(* IEC 61131-3 sources: moqui-plc/codesys-v4/moqui-plc.fbsdev/moqui.iecapp^/moqui/runtime/component/mantle-hvac/src/main/mantle/hvac, 3 files *)

(* ---- Main.fb.st ---- *)
(*
 * NOTE: In general, the Main component implements the control logic of automated industrial systems (Finite State Machine - FSM)
 * using hierarchical control architectures. It separates control policies from implementation mechanisms,
 * and diagnostic mechanisms from failure/error reaction and system reset policies.
*)

(* Example of a supervisor FSM for a civil HVAC air-handling unit (AHU).
 *
 * Topology:
 *   Mode A Thermostat cooling -> Cooling
 *   Mode B Cooling with RH% dehumidification -> Cooling  (rhControlEnabled=TRUE)
 *   Mode C Winter heating -> Heating
 *   Mode D Heating with RH% control -> Heating (rhControlEnabled=TRUE)
 *   Mode E Interval dehumidification (on/off) -> Drying
 *   Mode F Dehumidification by RH% target -> Drying (rhControlEnabled=TRUE)
 *
 * Output function - which device groups are enabled per state:
 *
 *   State          Cold Group   Hot Group   AHU Fan   Air Flow
 *   -
 *   Standby            OFF         OFF        OFF       OFF
 *   Ventilation        OFF         OFF        ON        ON
 *   Cooling            ON          OFF        ON        ON
 *   Heating            OFF         ON         ON        ON
 *   Drying             ON          ON         ON        ON
 *   Fault              OFF         OFF        OFF       OFF
 *
 * MainRuleEngine generates transition requests; Main consumes them.
 * DeviceManager orchestrates the individual device FBs.
 *
 * Call order in the PLC task:
 *   InputSignalUpdate -> Main -> DeviceManager -> OutputSignalUpdate
 *)
FUNCTION_BLOCK Main

	VAR_INPUT
		operationType : OperatingMode;
		enable : BOOL;
		deviceConfigContextResetRequest : BOOL := FALSE;
	END_VAR
	VAR_OUTPUT
		done : BOOL;
		error : BOOL;
	END_VAR
	VAR CONSTANT
		componentName : STRING := 'HVAC_DEMO_PLC';
	END_VAR
	VAR
		(* Logger facade *)
		logger : LoggerFacade;
		(* FSM transition logic *)
		ruleEngine : MainRuleEngine;
		(* Define a nested FSMs for managing air distribution subsystem. *)
		airDistribCtrl : AirDistributionController;
		(* HAL manager *)
		deviceManager : DeviceManager;
		(* Periodic logical-parameter logger *)
		logParameters : ParameterLogger;
		(* Previous status, so that the FSM state is logged on change only *)
		statusOld : MainStatus := MainStatus.Standby;
	END_VAR

	(* Logger facade init *)
	logger.enable := TRUE; logger.loggerName := componentName;

	IF NOT enable THEN RETURN; END_IF

	(* Init: device setup and configuration *)
	IF (operationType = operatingMode.Init) THEN
		logger(message := 'Setup and configuration of all devices.', level := LogLevel.DEBUG);
		(*
	     * The static device configuration parameters are mapped directly by the device config manager (recipe manager),
		 * while only the dynamic parameters are mapped below in the standby status.
		 *)
		(* Reset signal manager *)
		ec.dev.signalMgmt(operationType := SignalMgmtOperatingMode.Reset, loggerName := componentName);
		ec.dev.status := MainStatus.Standby;
		ec.dev.actualRuntime := 0;
		ec.dev.actualBreakDuration := 0;
		ec.dev.processActualDuration := 0;
		ec.dev.processRemainingDuration := 0;
		ec.dev.timeBreakEnabled := FALSE;
		ec.dev.isCompleted := FALSE;
		airDistribCtrl(operationType := OperatingMode.Init, enable := FALSE, clock1s := FALSE);
		done := FALSE;
	ELSIF deviceConfigContextResetRequest THEN
		logger(message := 'Reset HVAC device config context.', level := LogLevel.DEBUG);
		(*
	     * Lightweight reset between recipes: keep device init/homing in the Init path,
		 * but clear runtime state inherited from the previous device config.
	     *)
		ec.dev.status := MainStatus.Standby;
		ec.dev.lastStatus := MainStatus.Standby;
		ec.dev.actualRuntime := 0;
		ec.dev.actualBreakDuration := 0;
		ec.dev.processActualDuration := 0;
		ec.dev.processRemainingDuration := 0;
		ec.dev.timeBreakEnabled := FALSE;
		ec.dev.isCompleted := FALSE;
		airDistribCtrl(operationType := OperatingMode.Init, enable := FALSE, clock1s := FALSE);
		done := FALSE;
	ELSE
		(* FSM transition-condition rule engine *)
		ruleEngine(operationType := operationType);
	END_IF;

		(*
		 * Preserve the originating phase while idling in Standby so thermostat-driven
		 * Heating/Cooling recipes can stop/start repeatedly until isCompleted becomes TRUE.
		 * Init still stamps Standby, which keeps fresh-start logic for a newly loaded recipe.
		 * A temporary thermal override of Drying (Drying -> Cooling/Heating) keeps Drying as the
		 * originating phase: MainRuleEngine returns to Drying from Cooling/Heating while
		 * lastStatus = Drying, so it must stay Drying for the whole override, not for one scan.
	     *)
		IF operationType = OperatingMode.Init THEN
			ec.dev.lastStatus := ec.dev.status;
		ELSIF (ec.dev.status <> MainStatus.Standby)
				AND NOT ((ec.dev.lastStatus = MainStatus.Drying)
					AND ((ec.dev.status = MainStatus.Cooling) OR (ec.dev.status = MainStatus.Heating))) THEN
			ec.dev.lastStatus := ec.dev.status;
		END_IF;

	(* Fault overrides any other state *)
	IF ec.dev.faultRequest THEN ec.dev.status := MainStatus.Fault; END_IF;

	(* Main FSM - Output function + State-update function *)
	CASE ec.dev.status OF
	    (* Standby / Homing: all groups off, wait for the next phase request. *)
		MainStatus.Standby :
			ec.dev.standbyRequest := FALSE;

			(* FSM Output function - everything disabled *)
			ec.dev.coldGroupEnableRequest := FALSE;
			ec.dev.coldGroupDisableRequest := TRUE;
			ec.dev.hotGroupEnableRequest := FALSE;
			ec.dev.hotGroupDisableRequest := TRUE;
			ec.dev.ahuFanEnableRequest := FALSE;
			ec.dev.airFlowEnableRequest := FALSE;
			ec.dev.airFlowDisableRequest := TRUE;

			(* FSM status update function *)
			IF ec.dev.ventilationRequest THEN
				ec.dev.status := MainStatus.Ventilation;
			ELSIF ec.dev.coolingRequest THEN
				ec.dev.status := MainStatus.Cooling;
			ELSIF ec.dev.heatingRequest THEN
				ec.dev.status := MainStatus.Heating;
			ELSIF ec.dev.dryingRequest THEN
				ec.dev.status := MainStatus.Drying;
			END_IF;

	    (* Ventilation: AHU + air flow control only - no temperature conditioning. *)
		MainStatus.Ventilation :
			ec.dev.ventilationRequest := FALSE;

			(* FSM output function *)
			ec.dev.coldGroupEnableRequest := FALSE;
			ec.dev.coldGroupDisableRequest := TRUE;
			ec.dev.hotGroupEnableRequest := FALSE;
			ec.dev.hotGroupDisableRequest := TRUE;
			ec.dev.ahuFanEnableRequest := TRUE;
			ec.dev.airFlowEnableRequest := TRUE;
			ec.dev.airFlowDisableRequest := FALSE;

			(* FSM status update function *)
			IF ec.dev.standbyRequest THEN
				ec.dev.status := MainStatus.Standby;
			ELSIF ec.dev.coolingRequest THEN
				ec.dev.status := MainStatus.Cooling;
			ELSIF ec.dev.heatingRequest THEN
				ec.dev.status := MainStatus.Heating;
			ELSIF ec.dev.dryingRequest THEN
				ec.dev.status := MainStatus.Drying;
			END_IF;

	    (*
	     * Cooling: cold group + AHU + air flow control.
	     * Mode A (no RH ctrl) and Mode B (with RH dehumidification, rhControlEnabled=TRUE).
	     * In Mode B the hot group is also enabled to re-heat after dehumidification;
	     * that secondary enable is issued by MainRuleEngine via heatingRequest/dryingRequest
	     * transitions rather than here, keeping output function clean.
	     *)
		MainStatus.Cooling :
			ec.dev.coolingRequest := FALSE;

			(* FSM output function *)
			ec.dev.coldGroupEnableRequest := TRUE;
			ec.dev.coldGroupDisableRequest := FALSE;
			ec.dev.hotGroupEnableRequest := FALSE;
			ec.dev.hotGroupDisableRequest := TRUE;
			ec.dev.ahuFanEnableRequest := TRUE;
			ec.dev.airFlowEnableRequest := TRUE;
			ec.dev.airFlowDisableRequest := FALSE;

			(* FSM status update function *)
			IF ec.dev.standbyRequest THEN
				ec.dev.status := MainStatus.Standby;
			ELSIF ec.dev.dryingRequest THEN
				ec.dev.status := MainStatus.Drying;
			ELSIF ec.dev.ventilationRequest THEN
				ec.dev.status := MainStatus.Ventilation;
			END_IF;

	    (*
	     * Heating: hot group + AHU + air flow control.
	     * Mode C (no RH ctrl) and Mode D (with RH ctrl).
	     *)
		MainStatus.Heating :
			ec.dev.heatingRequest := FALSE;

			(* FSM output function *)
			ec.dev.coldGroupEnableRequest := FALSE;
			ec.dev.coldGroupDisableRequest := TRUE;
			ec.dev.hotGroupEnableRequest := TRUE;
			ec.dev.hotGroupDisableRequest := FALSE;
			ec.dev.ahuFanEnableRequest := TRUE;
			ec.dev.airFlowEnableRequest := TRUE;
			ec.dev.airFlowDisableRequest := FALSE;

			(* FSM status update function *)
			IF ec.dev.standbyRequest THEN
				ec.dev.status := MainStatus.Standby;
			ELSIF ec.dev.dryingRequest THEN
				ec.dev.status := MainStatus.Drying;
			ELSIF ec.dev.ventilationRequest THEN
				ec.dev.status := MainStatus.Ventilation;
			END_IF;

	    (*
	     * Drying: cold + hot + AHU + air flow control.
	     * Mode E (interval on/off) and Mode F (RH% controlled).
	     * During break the rule engine transitions to Standby; returns here
	     * when the break is complete.
	     *)
		MainStatus.Drying :
			ec.dev.dryingRequest := FALSE;

			(* FSM output function *)
			ec.dev.coldGroupEnableRequest := TRUE;
			ec.dev.coldGroupDisableRequest := FALSE;
			ec.dev.hotGroupEnableRequest := TRUE;
			ec.dev.hotGroupDisableRequest := FALSE;
			ec.dev.ahuFanEnableRequest := TRUE;
			ec.dev.airFlowEnableRequest := TRUE;
			ec.dev.airFlowDisableRequest := FALSE;

			(* FSM status update function *)
			IF ec.dev.standbyRequest THEN
				ec.dev.status := MainStatus.Standby;
			ELSIF ec.dev.heatingRequest THEN
				ec.dev.status := MainStatus.Heating;
			ELSIF ec.dev.coolingRequest THEN
				ec.dev.status := MainStatus.Cooling;
			ELSIF ec.dev.ventilationRequest THEN
				ec.dev.status := MainStatus.Ventilation;
			END_IF;

	    (* Fault: all groups off; wait for signal manager to clear all alarms. *)
		MainStatus.Fault :
			ec.dev.faultRequest := FALSE;

			(* FSM output function *)
			error := TRUE;
			ec.dev.coldGroupEnableRequest := FALSE;
			ec.dev.coldGroupDisableRequest := TRUE;
			ec.dev.hotGroupEnableRequest := FALSE;
			ec.dev.hotGroupDisableRequest := TRUE;
			ec.dev.ahuFanEnableRequest := FALSE;
			ec.dev.airFlowEnableRequest := FALSE;
			ec.dev.airFlowDisableRequest := TRUE;

			(* Return to Standby only when all alarms have been cleared *)
			IF (ec.dev.signalMgmt.cumulativeOutputAction = SignalOutputAction.None) THEN
				error := FALSE;
				ec.dev.status := MainStatus.Standby;
			END_IF;
	END_CASE;

	(*
	 * Air distribution is a subordinate subsystem:
	 * it runs only when the main FSM requests air flow and the recipe explicitly
	 * enables alternating high/low air distribution.
	 *)
	airDistribCtrl(
		operationType := operationType,
		enable := ec.dev.airFlowEnableRequest AND ec.dev.airDistributionEnabled,
		clock1s := ec.clks.clock1s);

	done := ec.dev.isCompleted;

	(* Log the FSM state on change only: a message every scan would fill the log buffer. *)
	IF ec.dev.status <> statusOld THEN
		CASE ec.dev.status OF
			MainStatus.Standby : logger(message := 'Standby.', level := LogLevel.Info);
			MainStatus.Ventilation : logger(message := 'Ventilation.', level := LogLevel.Info);
			MainStatus.Cooling : logger(message := 'Cooling.', level := LogLevel.Info);
			MainStatus.Heating : logger(message := 'Heating.', level := LogLevel.Info);
			MainStatus.Drying : logger(message := 'Drying.', level := LogLevel.Info);
			MainStatus.Fault : logger(message := 'Fault.', level := LogLevel.Error);
		END_CASE;
		statusOld := ec.dev.status;
	END_IF;

	(* Device orchestration (HAL) *)
	deviceManager(operationType := operationType);

	(* Log the coherent post-device-update parameter snapshot. *)
	logParameters(operationType := operationType);
	END_FUNCTION_BLOCK

(* ---- MainRuleEngine.fb.st ---- *)
(*
 * MainRuleEngine - transition-condition logic for the HVAC supervisor FSM.
 *
 * Responsibilities:
 *   1. Reset transition requests to safe defaults.
 *   2. Run the signal management engine (fault / alarm / warning detection).
 *   3. Compute boolean predicates from sensor feedback and recipe setpoints.
 *   4. Implement the per-state transition-condition rules.
 *
 * Default / persistence convention
 * At the top of every scan standbyRequest is set TRUE (safe default).
 * Each ACTIVE-state CASE block MUST:
 *   - Set standbyRequest := FALSE (keep current state) in the ELSE branch.
 *   - Set standbyRequest := TRUE (or leave as-is) when an EXIT condition is met.
 *   - Set standbyRequest := FALSE and another*Request := TRUE to switch phase.
 *
 * Without the ELSE branch the system would exit any active state to Standby
 * on the very first scan - a single-scan flash rather than a persistent phase.
 *
 * Operating modes:
 *   Mode A Thermostat Cooling -> Cooling
 *   Mode B Cooling with RH% dehumidification -> Cooling (rhControlEnabled)
 *   Mode C Winter Heating -> Heating
 *   Mode D Heating with RH% control -> Heating (rhControlEnabled)
 *   Mode E Interval Dehumidification (on/off) -> Drying <-> Standby (break)
 *   Mode F Dehumidification by RH% target -> Drying (rhControlEnabled)
 *
 * Duct safety (duct sensors):
 *   The duct T+RH sensor monitors supply-air conditions upstream of the zone.
 *   Limit violations raise alarms to protect equipment and occupants.
 *   ductTempOverMax -> supply air too hot -> ImmediateStop
 *   ductTempUnderMin -> supply air too cold -> ImmediateStop
 *   ductRhOverMax -> supply air saturated -> Warning only (condensation risk)
 *)
FUNCTION_BLOCK MainRuleEngine

	VAR_INPUT
		operationType : OperatingMode := OperatingMode.Run;
	END_VAR
	VAR_OUTPUT
		error : BOOL;
	END_VAR
	VAR
		(* Device diagnostics *)
		deviceDiags : DeviceDiagnostics;
	END_VAR

	(* Reset transition requests to safe defaults.
	 *
	 * standbyRequest = TRUE -> return to / stay in Standby (safe default).
	 * Active-state CASE blocks override to FALSE to keep the current phase alive,
	 * or set another *Request to switch phases.
	 *)
	ec.dev.faultRequest := FALSE;
	ec.dev.standbyRequest := TRUE;
	ec.dev.heatingRequest := FALSE;
	ec.dev.coolingRequest := FALSE;
	ec.dev.ventilationRequest := FALSE;
	ec.dev.dryingRequest := FALSE;

	deviceDiags(operationType := operationType, error => error);

	(* Compute sensor predicates *)

	(* Process temperature sensor *)
	ec.dev.tempInRange := (ec.dev.tempFeedback >= ec.dev.tempMin + ec.dev.tempHysteresis)
		AND (ec.dev.tempFeedback <= ec.dev.tempMax - ec.dev.tempHysteresis);
	ec.dev.tempAtSetpoint := ABS(ec.dev.tempFeedback - ec.dev.tempSetpoint) <= ec.dev.tempHysteresis;
	(* Normal thermostat thresholds are independent from the absolute alarm limits. *)
	ec.dev.tempAboveSetpointBand := ec.dev.tempFeedback >= (ec.dev.tempSetpoint + ec.dev.tempHysteresis);
	ec.dev.tempBelowSetpointBand := ec.dev.tempFeedback <= (ec.dev.tempSetpoint - ec.dev.tempHysteresis);
	ec.dev.tempOverMax := ec.dev.tempFeedback > ec.dev.tempMax;
	ec.dev.tempOverMin := ec.dev.tempFeedback > ec.dev.tempMin;
	ec.dev.tempUnderMin := ec.dev.tempFeedback < ec.dev.tempMin;
	ec.dev.tempUnderMax := ec.dev.tempFeedback < ec.dev.tempMax;

	(* Process RH sensor *)
	ec.dev.rhAtSetpoint := ABS(ec.dev.rhFeedback - ec.dev.rhSetpoint) <= ec.dev.rhHysteresis;
	ec.dev.rhOverMax := ec.dev.rhFeedback > ec.dev.rhMax - ec.dev.rhHysteresis;
	ec.dev.rhUnderMin := ec.dev.rhFeedback < ec.dev.rhMin + ec.dev.rhHysteresis;
	ec.dev.rhOverMin := ec.dev.rhFeedback > ec.dev.rhMin;
	ec.dev.rhUnderMax := ec.dev.rhFeedback < ec.dev.rhMax;

	(* Duct sensor - safety predicates *)
	ec.dev.ductTempOverMax := ec.dev.ductTempFeedback > ec.dev.ductTempMax;
	ec.dev.ductTempUnderMin := ec.dev.ductTempFeedback < ec.dev.ductTempMin;
	ec.dev.ductRhOverMax := ec.dev.ductRhFeedback > ec.dev.ductRhMax;

	(*
	 * Process timing - run / break cycle.
	 *
	 * processActualDuration must NOT advance while the FSM is in Standby
	 * waiting for a phase to start (i.e. not in a break).
	 * If it did, isCompleted could fire while the process has not yet begun,
	 * causing the phase to complete immediately without doing any work.
	 *
	 * Counting rules:
	 *   Break (timeBreakEnabled=TRUE, status=Standby): advance processActualDuration + actualBreakDuration.
	 *   Active (status != Standby): advance processActualDuration + actualRuntime.
	 *   Idle (status=Standby, NOT timeBreakEnabled): no counters advance.
	 *)
	IF ec.clks.clock1s THEN
		IF ec.dev.timeBreakEnabled AND ec.dev.status = MainStatus.Standby THEN
			(* Break counting *)
			ec.dev.processActualDuration := ec.dev.processActualDuration + 1;
			ec.dev.actualBreakDuration := ec.dev.actualBreakDuration + 1;
			IF ec.dev.estimatedBreakDuration > 0 THEN
				(* Break ends when both minimum and estimated durations are met; reset counters for next run *)
				IF (ec.dev.actualBreakDuration >= ec.dev.estimatedBreakDuration)
						AND (ec.dev.actualBreakDuration >= ec.dev.minBreakDuration) THEN
					ec.dev.timeBreakEnabled := FALSE;
					ec.dev.actualRuntime := 0;
					ec.dev.actualBreakDuration := 0;
				END_IF;
			END_IF;
		ELSIF ec.dev.status <> MainStatus.Standby THEN
			(* Active run counting - only while the FSM is in an active phase state *)
			ec.dev.processActualDuration := ec.dev.processActualDuration + 1;
			ec.dev.actualRuntime := ec.dev.actualRuntime + 1;
			IF ec.dev.estimatedRuntime > 0 THEN
				IF NOT ec.dev.timeBreakEnabled
						AND (ec.dev.actualRuntime >= ec.dev.estimatedRuntime)
						AND (ec.dev.actualRuntime >= ec.dev.minRuntime) THEN
					ec.dev.timeBreakEnabled := TRUE;
					ec.dev.actualBreakDuration := 0;
				END_IF;
			END_IF;
		ELSIF (ec.dev.lastStatus = MainStatus.Cooling OR ec.dev.lastStatus = MainStatus.Heating)
				AND NOT ec.dev.isCompleted THEN
			(* Thermostat dwell between active cycles counts toward phase duration,
			 * but does not count as active runtime. *)
			ec.dev.processActualDuration := ec.dev.processActualDuration + 1;
		END_IF;

		(* Remaining duration, saturated at zero: the durations are UDINT and a phase can outlast its estimate. *)
		IF ec.dev.processEstimatedDuration > ec.dev.processActualDuration THEN
			ec.dev.processRemainingDuration := ec.dev.processEstimatedDuration - ec.dev.processActualDuration;
		ELSE
			ec.dev.processRemainingDuration := 0;
		END_IF;

		(* isCompleted is independent of the run/break cycle:
		 * a phase with only processEstimatedDuration set (no run/break) must also complete. *)
		IF ec.dev.processEstimatedDuration > 0 THEN
			ec.dev.isCompleted :=
				(ec.dev.processActualDuration >= ec.dev.processEstimatedDuration)
				AND (ec.dev.processActualDuration >= ec.dev.processMinDuration);
		END_IF;
	END_IF;

	(* Fault gate *)
	IF error OR ((ec.dev.signalMgmt.cumulativeOutputAction AND SignalOutputAction.ImmediateStop) <> 0) THEN
		ec.dev.faultRequest := TRUE;
		RETURN;
	END_IF;

	(*
	 * Transition-condition rule engine
	 *
	 * Persistence rule: every active-state CASE MUST end with
	 *   ELSE dev.standbyRequest := FALSE; (* keep current state alive *)
	 * to prevent the scan-level default (standbyRequest=TRUE) from immediately
	 * bouncing the FSM back to Standby before the exit condition is reached.
	 *)
	CASE ec.dev.status OF
	    (*
	     * Standby - decide next phase.
	     * Default standbyRequest=TRUE keeps the system here.
	     * Override when an external condition requires re-entering a phase.
	     *)
		MainStatus.Standby :
			(*
			 * Transition-condition evaluation order:
			 *   1. Safety overrides (cooling/heating if temperature out of limits).
			 *   2. Phase-resume conditions (dehumidification after break).
			 *   3. Fresh-start dehumidification (new recipe loaded, lastStatus=Standby after Init).
			 *   4. Hold-in-Standby (isCompleted) - checked LAST.
			 *
			 * isCompleted is evaluated last so that phase-transition conditions are always
			 * reachable.  The guard dev.lastStatus=Standby in condition 3 makes it safe:
			 * that guard is only TRUE after Init has run (Init sets dev.status=Standby, so
			 * line-97 lastStatus:=status writes Standby), which also resets isCompleted=FALSE.
			 * In the one-scan gap between a phase exit (isCompleted=TRUE, lastStatus=Cooling/
			 * Drying/…) and Init, lastStatus != Standby, so condition 3 cannot fire, and
			 * condition 4 correctly holds the FSM in Standby until configMgmt advances.
			 *)
			IF (ec.dev.lastStatus = MainStatus.Cooling OR ec.dev.lastStatus = MainStatus.Standby)
					AND ec.dev.tempAboveSetpointBand THEN
				(* Temperature above the thermostat band -> start/resume cooling. *)
				ec.dev.standbyRequest := FALSE;
				ec.dev.coolingRequest := TRUE;

			ELSIF (ec.dev.lastStatus = MainStatus.Heating OR ec.dev.lastStatus = MainStatus.Standby)
					AND ec.dev.tempBelowSetpointBand THEN
				(* Temperature below the thermostat band -> start/resume heating. *)
				ec.dev.standbyRequest := FALSE;
				ec.dev.heatingRequest := TRUE;

			ELSIF ec.dev.lastStatus = MainStatus.Drying
					AND NOT ec.dev.timeBreakEnabled
					AND NOT ec.dev.isCompleted
					AND ec.dev.tempInRange
					AND (NOT ec.dev.rhControlOnly
					OR (ec.dev.rhControlEnabled AND ec.dev.rhOverMax)) THEN
				(*
				 * End of break: resume dehumidification run when all conditions are met:
				 *   - break elapsed (NOT timeBreakEnabled)
				 *   - process not yet complete (NOT isCompleted)
				 *   - temperature back in process window (tempInRange)
				 *   - humidity still needs treatment
				 *)
				ec.dev.standbyRequest := FALSE;
				ec.dev.dryingRequest := TRUE;

			ELSIF ec.dev.lastStatus = MainStatus.Standby
					AND NOT ec.dev.tempOverMax
					AND ec.dev.rhOverMax THEN
				(*
				 * Fresh dehumidification recipe loaded: start when temperature is safe (<= tempMax)
				 * and humidity needs treatment.
				 *
				 * NOT tempOverMax (instead of tempInRange) eliminates the dead zone at
				 * tempFeedback in (tempMax-hyst, tempMax] that would leave the FSM stuck in
				 * Standby after a cooling phase delivered temp near the top of the window.
				 * If temp is below tempMin the Drying state switches to Heating temporarily,
				 * then returns to Drying once tempOverMin.
				 *)
				ec.dev.standbyRequest := FALSE;
				ec.dev.dryingRequest := TRUE;

			ELSIF ec.dev.isCompleted THEN
				ec.dev.standbyRequest := TRUE; (* Explicit: work done, hold here until configMgmt advances *)

			(* No ELSE needed here: standbyRequest=TRUE default holds Standby *)
			END_IF;

	    (*
	     * Ventilation - AHU + air flow only.
	     * No automatic exit; operator or recipe change triggers Standby.
	     *)
		MainStatus.Ventilation :
			IF ec.dev.isCompleted THEN
				ec.dev.standbyRequest := TRUE;
			ELSE
				ec.dev.standbyRequest := FALSE; (* Keep ventilating *)
			END_IF;

	    (*
	     * Cooling - cold group + AHU.
	     * Mode A: thermostat-only (no RH control).
	     * Mode B: with RH dehumidification - when RH reaches setpoint switch to Drying.
	     *
	     * EXIT conditions (standbyRequest=TRUE):
	     *   tempBelowSetpointBand -> lower thermostat threshold reached.
	     *   isCompleted -> work-effort complete.
	     * SWITCH conditions (standbyRequest=FALSE):
	     *   lastStatus=Drying + tempUnderMax -> resume dehumidification.
	     * ELSE -> keep cooling (temperature still above tempMin).
	     *)
		MainStatus.Cooling :
			IF ec.dev.tempBelowSetpointBand OR ec.dev.isCompleted THEN
				ec.dev.standbyRequest := TRUE;
			ELSIF ec.dev.lastStatus = MainStatus.Drying
					AND (ec.dev.tempUnderMax
					OR (ec.dev.rhControlEnabled AND ec.dev.rhOverMax AND ec.dev.tempUnderMax)) THEN
				ec.dev.standbyRequest := FALSE;
				ec.dev.dryingRequest := TRUE;
			ELSE
				ec.dev.standbyRequest := FALSE; (* Keep cooling - tempFeedback still above tempMin *)
			END_IF;

	    (*
	     * Heating - hot group + AHU.
	     * Mode C (no RH ctrl) / Mode D (with RH ctrl).
	     *
	     * EXIT: upper thermostat threshold reached or isCompleted.
	     * SWITCH to Drying: temperature restored to process window.
	     * ELSE: keep heating.
	     *)
		MainStatus.Heating :
			IF ec.dev.isCompleted OR ec.dev.tempAboveSetpointBand THEN
				ec.dev.standbyRequest := TRUE;
			ELSIF (ec.dev.lastStatus = MainStatus.Drying AND ec.dev.tempOverMin)
					OR (ec.dev.rhControlEnabled AND ec.dev.rhOverMax) THEN
				ec.dev.standbyRequest := FALSE;
				ec.dev.dryingRequest  := TRUE;
			ELSE
				ec.dev.standbyRequest := FALSE; (* Keep heating - tempFeedback still below tempMax *)
			END_IF;

	    (*
	     * Drying - cold + hot + AHU (Mode E / Mode F).
	     *
	     * Normal end conditions:
	     *   Time-based (!rhControlOnly): T in range AND runtime elapsed.
	     *   RH-only: RH <= rhMin AND minimum runtime elapsed.
	     *   RH+time: RH <= rhMin (timer managed externally).
	     *   isCompleted: work-effort done.
	     * Break trigger: timeBreakEnabled -> Standby (returns here after break).
	     * Override to Cooling: tempOverMax.
	     * Override to Heating: tempUnderMin.
	     * ELSE: keep dehumidifying.
	     *)
		MainStatus.Drying :
			IF ec.dev.isCompleted THEN
				ec.dev.standbyRequest := TRUE;
			ELSIF NOT ec.dev.rhControlOnly
					AND ec.dev.tempInRange
					AND (ec.dev.estimatedRuntime > 0)
					AND (ec.dev.actualRuntime > ec.dev.estimatedRuntime) THEN
				ec.dev.standbyRequest := TRUE; (* Time-based running completed *)
			ELSIF ec.dev.rhControlOnly
					AND ec.dev.rhUnderMin
					AND (ec.dev.actualRuntime >= ec.dev.minRuntime) THEN
				ec.dev.standbyRequest := TRUE; (* RH-only target reached *)
			ELSIF ec.dev.rhControlEnabled AND ec.dev.rhUnderMin THEN
				ec.dev.standbyRequest := TRUE; (* RH+time: humidity at minimum *)
			ELSIF ec.dev.timeBreakEnabled THEN
				ec.dev.standbyRequest := TRUE; (* Begin break - rule engine resumes Drying after break *)
			ELSIF ec.dev.tempOverMax THEN
				ec.dev.standbyRequest := FALSE;
				ec.dev.coolingRequest := TRUE;  (* Temporary cooling override *)
			ELSIF ec.dev.tempUnderMin THEN
				ec.dev.standbyRequest := FALSE;
				ec.dev.heatingRequest := TRUE;  (* Temporary heating override *)
			ELSE
				ec.dev.standbyRequest := FALSE; (* Keep dehumidifying - process ongoing *)
			END_IF;
	END_CASE;
	END_FUNCTION_BLOCK

(* ---- ParameterLogger.fb.st ---- *)
(*
 * Periodic logger for the numeric parameters of the HVAC Application.
 *
 * Physical signal logging belongs to InputSignalUpdate and OutputSignalUpdate.
 * This block logs the logical values exposed through DeviceFacade. The source
 * of each event is the exact moqui.math.Parameter.parameterId from
	 * HVACDemoData.xml; loggerName is the owning Device.deviceId.
 *)
FUNCTION_BLOCK ParameterLogger

	VAR_INPUT
		operationType : OperatingMode;
	END_VAR
	VAR
		logger : LoggerFacade;
	END_VAR
	VAR CONSTANT
		componentName : STRING := 'HVAC_DEMO_PLC';
	END_VAR

	(* Log only one snapshot per minute, independently of the PLC task cycle. *)
	IF (operationType <> OperatingMode.Run) OR NOT ec.clks.clock1minute THEN RETURN; END_IF;

	logger.enable := TRUE;
	logger.loggerName := componentName;
	logger.payloadType := LogPayloadType.Numeric;
	logger.level := LogLevel.Info;
	(* The snapshot is a bounded burst of 29 events once a minute: not subject to the rate limit *)
	logger.maxEventsPerWindow := 0;

	(* Process setpoints and limits. *)
	logger(source := 'HvacTempSetpoint', numericValue := TO_LREAL(ec.dev.tempSetpoint));
	logger(source := 'HvacTempHysteresis', numericValue := TO_LREAL(ec.dev.tempHysteresis));
	logger(source := 'HvacTempMin', numericValue := TO_LREAL(ec.dev.tempMin));
	logger(source := 'HvacTempMax', numericValue := TO_LREAL(ec.dev.tempMax));
	logger(source := 'HvacRhSetpoint', numericValue := TO_LREAL(ec.dev.rhSetpoint));
	logger(source := 'HvacRhHysteresis', numericValue := TO_LREAL(ec.dev.rhHysteresis));
	logger(source := 'HvacRhMin', numericValue := TO_LREAL(ec.dev.rhMin));
	logger(source := 'HvacRhMax', numericValue := TO_LREAL(ec.dev.rhMax));
	logger(source := 'HvacDuctTempMin', numericValue := TO_LREAL(ec.dev.ductTempMin));
	logger(source := 'HvacDuctTempMax', numericValue := TO_LREAL(ec.dev.ductTempMax));
	logger(source := 'HvacDuctRhMax', numericValue := TO_LREAL(ec.dev.ductRhMax));

	(* Application timing parameters and runtime counters. *)
	logger(source := 'HvacSetPointTimeHigh', numericValue := TO_LREAL(ec.dev.setPointTimeHigh));
	logger(source := 'HvacSetPointTimeLow', numericValue := TO_LREAL(ec.dev.setPointTimeLow));
	logger(source := 'HvacEstimatedRuntime', numericValue := TO_LREAL(ec.dev.estimatedRuntime));
	logger(source := 'HvacMinRuntime', numericValue := TO_LREAL(ec.dev.minRuntime));
	logger(source := 'HvacEstimatedBreakDuration', numericValue := TO_LREAL(ec.dev.estimatedBreakDuration));
	logger(source := 'HvacMinBreakDuration', numericValue := TO_LREAL(ec.dev.minBreakDuration));
	logger(source := 'HvacProcessEstimatedDuration', numericValue := TO_LREAL(ec.dev.processEstimatedDuration));
	logger(source := 'HvacProcessMinDuration', numericValue := TO_LREAL(ec.dev.processMinDuration));
	logger(source := 'HvacProcessRemainingDuration', numericValue := TO_LREAL(ec.dev.processRemainingDuration));
	logger(source := 'HvacProcessActualDuration', numericValue := TO_LREAL(ec.dev.processActualDuration));
	logger(source := 'HvacActualRuntime', numericValue := TO_LREAL(ec.dev.actualRuntime));
	logger(source := 'HvacActualBreakDuration', numericValue := TO_LREAL(ec.dev.actualBreakDuration));

	(* Numeric machine references. *)
	logger(source := 'HvacAhuFanSpeedSetpoint', numericValue := TO_LREAL(ec.dev.ahuFanSpeedSetpoint));
	logger(source := 'HvacAirFlowRef', numericValue := TO_LREAL(ec.dev.airFlowRef));

	(* Process measurements. *)
	logger(source := 'HvacTempFeedback', numericValue := TO_LREAL(ec.dev.tempFeedback));
	logger(source := 'HvacRhFeedback', numericValue := TO_LREAL(ec.dev.rhFeedback));
	logger(source := 'HvacDuctTempFeedback', numericValue := TO_LREAL(ec.dev.ductTempFeedback));
	logger(source := 'HvacDuctRhFeedback', numericValue := TO_LREAL(ec.dev.ductRhFeedback));
	END_FUNCTION_BLOCK
